(* IEC 61131-3 sources: ZPLC/packages/zplc-ide/projects/conveyor_01_starter/src, 1 file *)

(* ---- Conveyor.st ---- *)
PROGRAM Conveyor

VAR_INPUT
    Start AT %I0.0 : BOOL;
    Stop AT %I0.1 : BOOL;
    Reset AT %I0.2 : BOOL;
    PartAtClassifier AT %I0.3 : BOOL;
    MetalDetected AT %I0.4 : BOOL;
    PartAtDiverter AT %I0.5 : BOOL;
    JamDetected AT %I0.6 : BOOL;
END_VAR

VAR
    Requested : BOOL := FALSE;
    MetalLatched : BOOL := FALSE;
END_VAR

VAR_OUTPUT
    BeltCommand AT %Q0.0 : BOOL;
    DiverterCommand AT %Q0.1 : BOOL;
    FaultLamp AT %Q0.2 : BOOL;
END_VAR

(* Educational host exercise: this incomplete starter intentionally omits the jam lockout.
   Lesson 4: stop the belt and light FaultLamp while JamDetected. Lesson 9: also latch the fault,
   release it only with Reset once the jam has cleared, and do not restart the belt without a new Start.
   Outputs still default FALSE on reset; never use this program on hardware. *)
IF Stop THEN
    Requested := FALSE;
ELSIF Start THEN
    Requested := TRUE;
END_IF;

IF PartAtClassifier AND MetalDetected THEN
    MetalLatched := TRUE;
END_IF;

BeltCommand := Requested;
DiverterCommand := BeltCommand AND PartAtDiverter AND MetalLatched;
FaultLamp := JamDetected;

IF PartAtDiverter OR Stop OR Reset THEN
    MetalLatched := FALSE;
END_IF;

END_PROGRAM
